Fanuc KAREL source: KT00217.KL

PROGRAM KT00217
%NOLOCKGROUP
VAR
  H1: ARRAY[2] OF SHORT
  B2: BOOLEAN
  OUT: BOOLEAN
BEGIN
  H1[1] = 2
    B2 = FALSE
  OUT = H1[1] AND B2
END KT00217
